// TIA Portal V21 export
FUNCTION_BLOCK "FB_Doser"   // FB6, SCL
// stored: Access Published, MemoryReserve 100, Namespace Dosing, SetENOAutomatically false
   VAR_INPUT
      Start : Bool;   // Start dosing
      Stop : Bool;   // Stop dosing
   END_VAR
   VAR_OUTPUT
      Dosing : Bool;   // Dosing is running
      Done : Bool;   // Dosing finished
   END_VAR
   VAR
      Filler { S7_SetPoint := 'True'} : "Filling.FB_Filler";   // Filler of the unit Filling
      Recipe { S7_SetPoint := 'True'} : "Filling.UDT_FillRecipe";   // Recipe of the unit Filling
   END_VAR
BEGIN

       REGION Dosing through the filler
           #Recipe.TargetVolume := 0.5;
           #Filler(Start := #Start, Stop := #Stop, Recipe := #Recipe);
           #Dosing := #Filler.Filling;
           #Done := #Filler.Done;
       END_REGION
END_FUNCTION_BLOCK
